(*
SPDX-FileCopyrightText: c 2026 Oleksandr Tiutyk <trofimich@gmail.com>
SPDX-License-Identifier: MIT
License: https://opensource.org/license/mit
*)

(*!
<summary>Groups fixed-capacity byte-list operations and overflow handling.</summary>
<description>
Owns the independent child instances and their fixed registration array. Use from one PLC task at a stable address.
</description>
*)

{attribute 'no_assign'}
{attribute 'no_explicit_call' := 'do not call this function block directly'}
FUNCTION_BLOCK StaticByteListTestGroup EXTENDS TOF_Testing.TestGroup<7>
VAR_STAT
	{attribute 'hide'}
	_ClassName : STRING := __POUNAME();
END_VAR
VAR
	_LoadFromAny : ByteListLoadFromAnyTest(name := "LoadFromAny", parent := THIS^, useDynamicStorage := FALSE);
	_GetAndSet : ByteListIndexedAccessTest(name := "GetAndSet", parent := THIS^, useDynamicStorage := FALSE);
	_Find : ByteListFindTest(name := "Find", parent := THIS^, useDynamicStorage := FALSE);
	_Remove : ByteListRemoveValueTest(name := "Remove", parent := THIS^, useDynamicStorage := FALSE);
	_RemoveAt : ByteListRemoveRangeTest(name := "RemoveAt", parent := THIS^, useDynamicStorage := FALSE);
	_Clear : ByteListClearTest(name := "Clear", parent := THIS^, useDynamicStorage := FALSE);
	_Overflow : StaticByteListOverflowTest(name := "Overflow", parent := THIS^);

	_Children : ARRAY [0.._ChildCount - 1] OF TOF_Testing.ITestElement :=
	[
		_LoadFromAny,
		_GetAndSet,
		_Find,
		_Remove,
		_RemoveAt,
		_Clear,
		_Overflow
	];
END_VAR

//! <summary>Borrows the fixed child array. Callers must not modify it.</summary>
{attribute 'monitoring' := 'call'}
PROPERTY Children : REFERENCE TO ARRAY [0.._ChildCount - 1] OF TOF_Testing.ITestElement
GET
Children REF= _Children;
END_GET
END_PROPERTY

//! <summary>Borrows the concrete class name. Callers must not modify it.</summary>
{attribute 'monitoring' := 'call'}
PROPERTY ClassName : REFERENCE TO STRING
GET
ClassName REF= _ClassName;
END_GET
END_PROPERTY

//! <summary>Borrows the compiler-initialized namespace name. Callers must not modify it.</summary>
{attribute 'monitoring' := 'call'}
PROPERTY NamespaceName : REFERENCE TO STRING
GET
NamespaceName REF= CurrentNamespace.Name;
END_GET
END_PROPERTY

//! <summary>Reports the concrete instance size in bytes.</summary>
{attribute 'monitoring' := 'call'}
PROPERTY SelfSize : ULINT
GET
SelfSize := XSIZEOF(THIS^);
END_GET
END_PROPERTY

END_FUNCTION_BLOCK

(* stored: Version 1.1.0.1
   POU StaticByteListTestGroup: Id {94c80802-b3f8-43a9-bdaa-a0d4f809151d}, SpecialFunc None
   Property Children: Id {3ae67d00-b05f-4c9c-8b9b-16dc6e1ed6cd}
   Get Get: Id {803e49c3-be78-416d-b30b-278a8e6fc51d}
   Property ClassName: Id {ada866b6-9be8-4f0d-b3aa-bf513ade245a}
   Get Get: Id {10318d7d-1a67-472f-aa2c-de1b9db97933}
   Property NamespaceName: Id {c70437a2-0697-4f34-818f-3330d47a7c3d}
   Get Get: Id {574a8d25-eae0-4889-a3bc-ed4489225b33}
   Property SelfSize: Id {c32ca8af-be97-4ba4-80c6-717a23c29332}
   Get Get: Id {01f9f3f0-90bf-4df3-b53d-179cb6563414} *)
